// Mitsubishi GX Works2 project: 2024.06.20   PLC: Q03UDV

PROGRAM MAIN
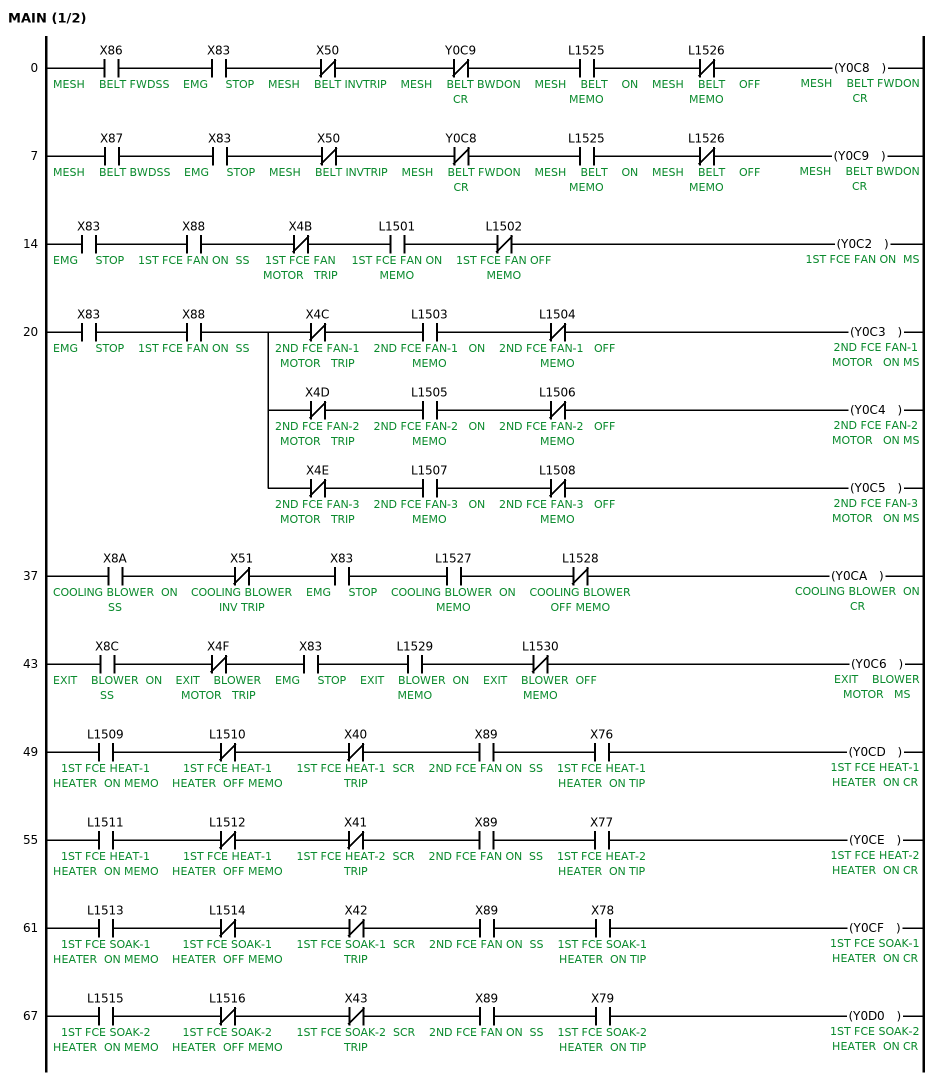
0     LD      X86  ; MESH    BELT FWDSS
      AND     X83  ; EMG     STOP
      ANI     X50  ; MESH    BELT INVTRIP
      ANI     Y0C9  ; MESH    BELT BWDON CR
      AND     L1525  ; MESH    BELT    ON MEMO
      ANI     L1526  ; MESH    BELT    OFF MEMO
      OUT     Y0C8  ; MESH    BELT FWDON CR
7     LD      X87  ; MESH    BELT BWDSS
      AND     X83  ; EMG     STOP
      ANI     X50  ; MESH    BELT INVTRIP
      ANI     Y0C8  ; MESH    BELT FWDON CR
      AND     L1525  ; MESH    BELT    ON MEMO
      ANI     L1526  ; MESH    BELT    OFF MEMO
      OUT     Y0C9  ; MESH    BELT BWDON CR
14    LD      X83  ; EMG     STOP
      AND     X88  ; 1ST FCE FAN ON  SS
      ANI     X4B  ; 1ST FCE FAN     MOTOR   TRIP
      AND     L1501  ; 1ST FCE FAN ON  MEMO
      ANI     L1502  ; 1ST FCE FAN OFF MEMO
      OUT     Y0C2  ; 1ST FCE FAN ON  MS
20    LD      X83  ; EMG     STOP
      AND     X88  ; 1ST FCE FAN ON  SS
      MPS
      ANI     X4C  ; 2ND FCE FAN-1   MOTOR   TRIP
      AND     L1503  ; 2ND FCE FAN-1   ON MEMO
      ANI     L1504  ; 2ND FCE FAN-1   OFF MEMO
      OUT     Y0C3  ; 2ND FCE FAN-1   MOTOR   ON MS
      MRD
      ANI     X4D  ; 2ND FCE FAN-2   MOTOR   TRIP
      AND     L1505  ; 2ND FCE FAN-2   ON MEMO
      ANI     L1506  ; 2ND FCE FAN-2   OFF MEMO
      OUT     Y0C4  ; 2ND FCE FAN-2   MOTOR   ON MS
      MPP
      ANI     X4E  ; 2ND FCE FAN-3   MOTOR   TRIP
      AND     L1507  ; 2ND FCE FAN-3   ON MEMO
      ANI     L1508  ; 2ND FCE FAN-3   OFF MEMO
      OUT     Y0C5  ; 2ND FCE FAN-3   MOTOR   ON MS
37    LD      X8A  ; COOLING BLOWER  ON SS
      ANI     X51  ; COOLING BLOWER  INV TRIP
      AND     X83  ; EMG     STOP
      AND     L1527  ; COOLING BLOWER  ON MEMO
      ANI     L1528  ; COOLING BLOWER  OFF MEMO
      OUT     Y0CA  ; COOLING BLOWER  ON CR
43    LD      X8C  ; EXIT    BLOWER  ON SS
      ANI     X4F  ; EXIT    BLOWER  MOTOR   TRIP
      AND     X83  ; EMG     STOP
      AND     L1529  ; EXIT    BLOWER  ON MEMO
      ANI     L1530  ; EXIT    BLOWER  OFF MEMO
      OUT     Y0C6  ; EXIT    BLOWER  MOTOR   MS
49    LD      L1509  ; 1ST FCE HEAT-1  HEATER  ON MEMO
      ANI     L1510  ; 1ST FCE HEAT-1  HEATER  OFF MEMO
      ANI     X40  ; 1ST FCE HEAT-1  SCR TRIP
      AND     X89  ; 2ND FCE FAN ON  SS
      AND     X76  ; 1ST FCE HEAT-1  HEATER  ON TIP
      OUT     Y0CD  ; 1ST FCE HEAT-1  HEATER  ON CR
55    LD      L1511  ; 1ST FCE HEAT-1  HEATER  ON MEMO
      ANI     L1512  ; 1ST FCE HEAT-1  HEATER  OFF MEMO
      ANI     X41  ; 1ST FCE HEAT-2  SCR TRIP
      AND     X89  ; 2ND FCE FAN ON  SS
      AND     X77  ; 1ST FCE HEAT-2  HEATER  ON TIP
      OUT     Y0CE  ; 1ST FCE HEAT-2  HEATER  ON CR
61    LD      L1513  ; 1ST FCE SOAK-1  HEATER  ON MEMO
      ANI     L1514  ; 1ST FCE SOAK-1  HEATER  OFF MEMO
      ANI     X42  ; 1ST FCE SOAK-1  SCR TRIP
      AND     X89  ; 2ND FCE FAN ON  SS
      AND     X78  ; 1ST FCE SOAK-1  HEATER  ON TIP
      OUT     Y0CF  ; 1ST FCE SOAK-1  HEATER  ON CR
67    LD      L1515  ; 1ST FCE SOAK-2  HEATER  ON MEMO
      ANI     L1516  ; 1ST FCE SOAK-2  HEATER  OFF MEMO
      ANI     X43  ; 1ST FCE SOAK-2  SCR TRIP
      AND     X89  ; 2ND FCE FAN ON  SS
      AND     X79  ; 1ST FCE SOAK-2  HEATER  ON TIP
      OUT     Y0D0  ; 1ST FCE SOAK-2  HEATER  ON CR
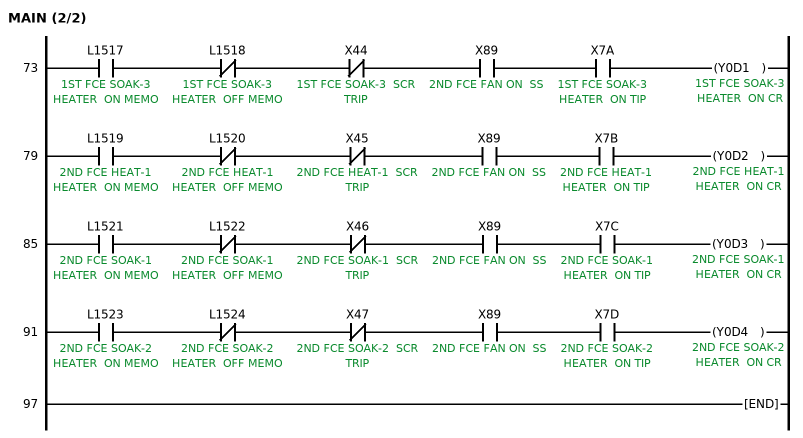
73    LD      L1517  ; 1ST FCE SOAK-3  HEATER  ON MEMO
      ANI     L1518  ; 1ST FCE SOAK-3  HEATER  OFF MEMO
      ANI     X44  ; 1ST FCE SOAK-3  SCR TRIP
      AND     X89  ; 2ND FCE FAN ON  SS
      AND     X7A  ; 1ST FCE SOAK-3  HEATER  ON TIP
      OUT     Y0D1  ; 1ST FCE SOAK-3  HEATER  ON CR
79    LD      L1519  ; 2ND FCE HEAT-1  HEATER  ON MEMO
      ANI     L1520  ; 2ND FCE HEAT-1  HEATER  OFF MEMO
      ANI     X45  ; 2ND FCE HEAT-1  SCR TRIP
      AND     X89  ; 2ND FCE FAN ON  SS
      AND     X7B  ; 2ND FCE HEAT-1  HEATER  ON TIP
      OUT     Y0D2  ; 2ND FCE HEAT-1  HEATER  ON CR
85    LD      L1521  ; 2ND FCE SOAK-1  HEATER  ON MEMO
      ANI     L1522  ; 2ND FCE SOAK-1  HEATER  OFF MEMO
      ANI     X46  ; 2ND FCE SOAK-1  SCR TRIP
      AND     X89  ; 2ND FCE FAN ON  SS
      AND     X7C  ; 2ND FCE SOAK-1  HEATER  ON TIP
      OUT     Y0D3  ; 2ND FCE SOAK-1  HEATER  ON CR
91    LD      L1523  ; 2ND FCE SOAK-2  HEATER  ON MEMO
      ANI     L1524  ; 2ND FCE SOAK-2  HEATER  OFF MEMO
      ANI     X47  ; 2ND FCE SOAK-2  SCR TRIP
      AND     X89  ; 2ND FCE FAN ON  SS
      AND     X7D  ; 2ND FCE SOAK-2  HEATER  ON TIP
      OUT     Y0D4  ; 2ND FCE SOAK-2  HEATER  ON CR
97    END
END_PROGRAM

PROGRAM HMI
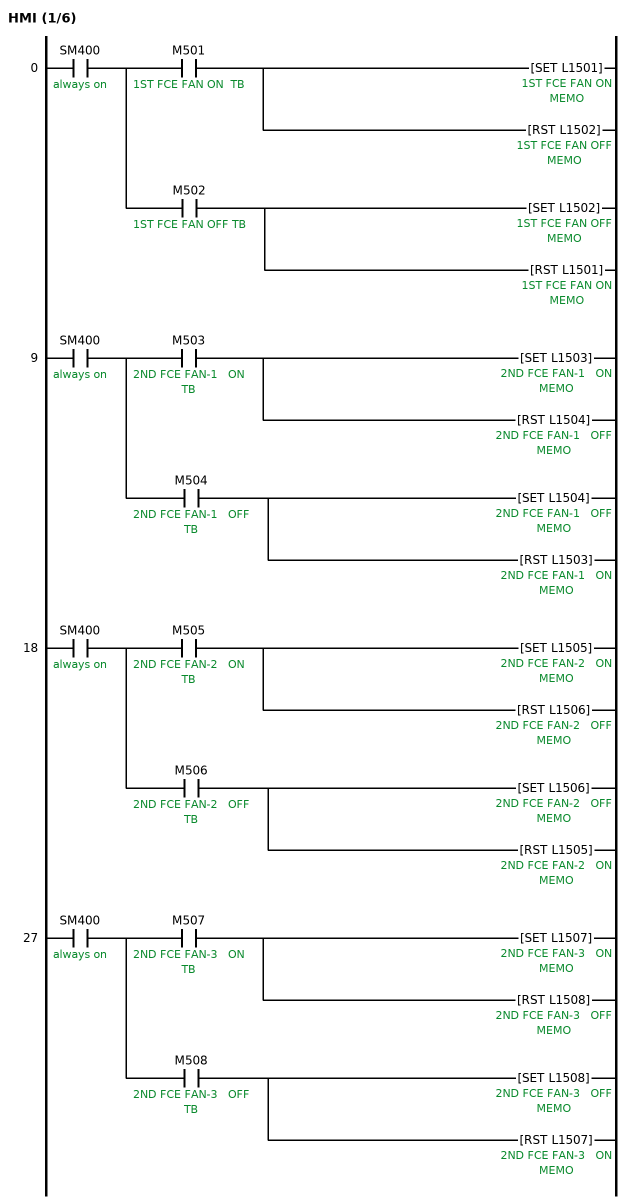
0     LD      SM400  ; always on
      MPS
      AND     M501  ; 1ST FCE FAN ON  TB
      SET     L1501  ; 1ST FCE FAN ON  MEMO
      RST     L1502  ; 1ST FCE FAN OFF MEMO
      MPP
      AND     M502  ; 1ST FCE FAN OFF TB
      SET     L1502  ; 1ST FCE FAN OFF MEMO
      RST     L1501  ; 1ST FCE FAN ON  MEMO
9     LD      SM400  ; always on
      MPS
      AND     M503  ; 2ND FCE FAN-1   ON TB
      SET     L1503  ; 2ND FCE FAN-1   ON MEMO
      RST     L1504  ; 2ND FCE FAN-1   OFF MEMO
      MPP
      AND     M504  ; 2ND FCE FAN-1   OFF TB
      SET     L1504  ; 2ND FCE FAN-1   OFF MEMO
      RST     L1503  ; 2ND FCE FAN-1   ON MEMO
18    LD      SM400  ; always on
      MPS
      AND     M505  ; 2ND FCE FAN-2   ON TB
      SET     L1505  ; 2ND FCE FAN-2   ON MEMO
      RST     L1506  ; 2ND FCE FAN-2   OFF MEMO
      MPP
      AND     M506  ; 2ND FCE FAN-2   OFF TB
      SET     L1506  ; 2ND FCE FAN-2   OFF MEMO
      RST     L1505  ; 2ND FCE FAN-2   ON MEMO
27    LD      SM400  ; always on
      MPS
      AND     M507  ; 2ND FCE FAN-3   ON TB
      SET     L1507  ; 2ND FCE FAN-3   ON MEMO
      RST     L1508  ; 2ND FCE FAN-3   OFF MEMO
      MPP
      AND     M508  ; 2ND FCE FAN-3   OFF TB
      SET     L1508  ; 2ND FCE FAN-3   OFF MEMO
      RST     L1507  ; 2ND FCE FAN-3   ON MEMO
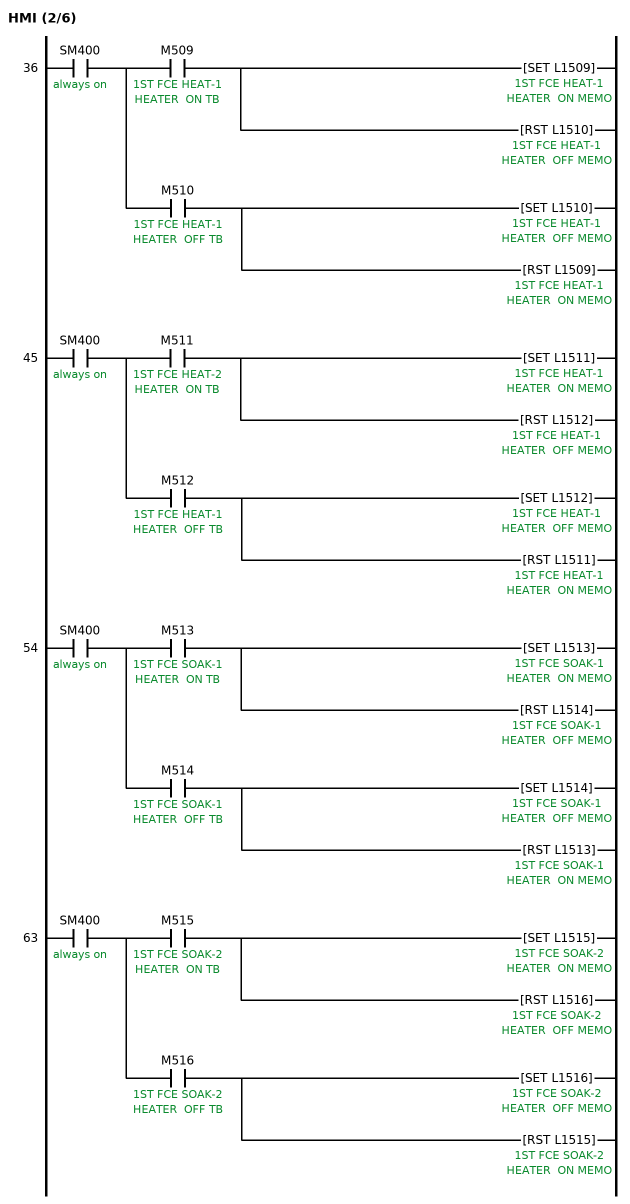
36    LD      SM400  ; always on
      MPS
      AND     M509  ; 1ST FCE HEAT-1  HEATER  ON TB
      SET     L1509  ; 1ST FCE HEAT-1  HEATER  ON MEMO
      RST     L1510  ; 1ST FCE HEAT-1  HEATER  OFF MEMO
      MPP
      AND     M510  ; 1ST FCE HEAT-1  HEATER  OFF TB
      SET     L1510  ; 1ST FCE HEAT-1  HEATER  OFF MEMO
      RST     L1509  ; 1ST FCE HEAT-1  HEATER  ON MEMO
45    LD      SM400  ; always on
      MPS
      AND     M511  ; 1ST FCE HEAT-2  HEATER  ON TB
      SET     L1511  ; 1ST FCE HEAT-1  HEATER  ON MEMO
      RST     L1512  ; 1ST FCE HEAT-1  HEATER  OFF MEMO
      MPP
      AND     M512  ; 1ST FCE HEAT-1  HEATER  OFF TB
      SET     L1512  ; 1ST FCE HEAT-1  HEATER  OFF MEMO
      RST     L1511  ; 1ST FCE HEAT-1  HEATER  ON MEMO
54    LD      SM400  ; always on
      MPS
      AND     M513  ; 1ST FCE SOAK-1  HEATER  ON TB
      SET     L1513  ; 1ST FCE SOAK-1  HEATER  ON MEMO
      RST     L1514  ; 1ST FCE SOAK-1  HEATER  OFF MEMO
      MPP
      AND     M514  ; 1ST FCE SOAK-1  HEATER  OFF TB
      SET     L1514  ; 1ST FCE SOAK-1  HEATER  OFF MEMO
      RST     L1513  ; 1ST FCE SOAK-1  HEATER  ON MEMO
63    LD      SM400  ; always on
      MPS
      AND     M515  ; 1ST FCE SOAK-2  HEATER  ON TB
      SET     L1515  ; 1ST FCE SOAK-2  HEATER  ON MEMO
      RST     L1516  ; 1ST FCE SOAK-2  HEATER  OFF MEMO
      MPP
      AND     M516  ; 1ST FCE SOAK-2  HEATER  OFF TB
      SET     L1516  ; 1ST FCE SOAK-2  HEATER  OFF MEMO
      RST     L1515  ; 1ST FCE SOAK-2  HEATER  ON MEMO
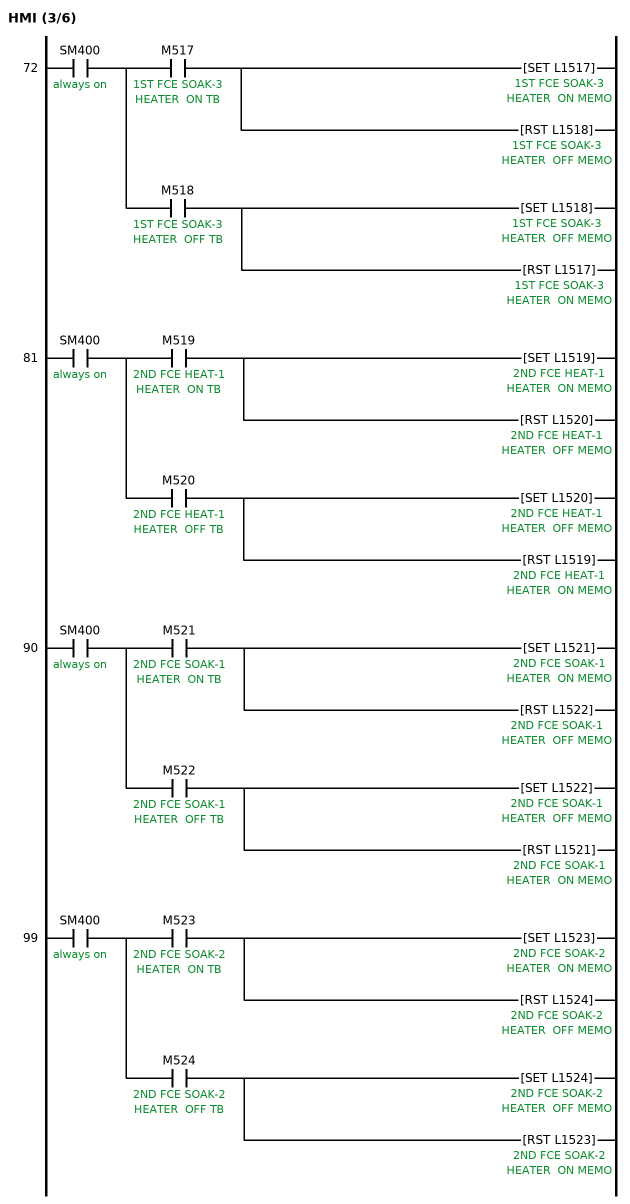
72    LD      SM400  ; always on
      MPS
      AND     M517  ; 1ST FCE SOAK-3  HEATER  ON TB
      SET     L1517  ; 1ST FCE SOAK-3  HEATER  ON MEMO
      RST     L1518  ; 1ST FCE SOAK-3  HEATER  OFF MEMO
      MPP
      AND     M518  ; 1ST FCE SOAK-3  HEATER  OFF TB
      SET     L1518  ; 1ST FCE SOAK-3  HEATER  OFF MEMO
      RST     L1517  ; 1ST FCE SOAK-3  HEATER  ON MEMO
81    LD      SM400  ; always on
      MPS
      AND     M519  ; 2ND FCE HEAT-1  HEATER  ON TB
      SET     L1519  ; 2ND FCE HEAT-1  HEATER  ON MEMO
      RST     L1520  ; 2ND FCE HEAT-1  HEATER  OFF MEMO
      MPP
      AND     M520  ; 2ND FCE HEAT-1  HEATER  OFF TB
      SET     L1520  ; 2ND FCE HEAT-1  HEATER  OFF MEMO
      RST     L1519  ; 2ND FCE HEAT-1  HEATER  ON MEMO
90    LD      SM400  ; always on
      MPS
      AND     M521  ; 2ND FCE SOAK-1  HEATER  ON TB
      SET     L1521  ; 2ND FCE SOAK-1  HEATER  ON MEMO
      RST     L1522  ; 2ND FCE SOAK-1  HEATER  OFF MEMO
      MPP
      AND     M522  ; 2ND FCE SOAK-1  HEATER  OFF TB
      SET     L1522  ; 2ND FCE SOAK-1  HEATER  OFF MEMO
      RST     L1521  ; 2ND FCE SOAK-1  HEATER  ON MEMO
99    LD      SM400  ; always on
      MPS
      AND     M523  ; 2ND FCE SOAK-2  HEATER  ON TB
      SET     L1523  ; 2ND FCE SOAK-2  HEATER  ON MEMO
      RST     L1524  ; 2ND FCE SOAK-2  HEATER  OFF MEMO
      MPP
      AND     M524  ; 2ND FCE SOAK-2  HEATER  OFF TB
      SET     L1524  ; 2ND FCE SOAK-2  HEATER  OFF MEMO
      RST     L1523  ; 2ND FCE SOAK-2  HEATER  ON MEMO
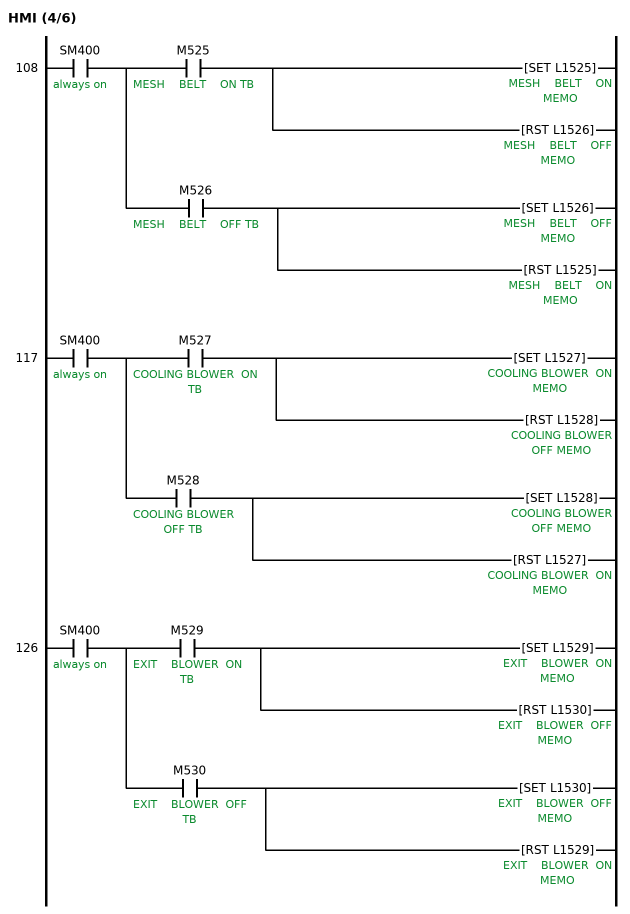
108   LD      SM400  ; always on
      MPS
      AND     M525  ; MESH    BELT    ON TB
      SET     L1525  ; MESH    BELT    ON MEMO
      RST     L1526  ; MESH    BELT    OFF MEMO
      MPP
      AND     M526  ; MESH    BELT    OFF TB
      SET     L1526  ; MESH    BELT    OFF MEMO
      RST     L1525  ; MESH    BELT    ON MEMO
117   LD      SM400  ; always on
      MPS
      AND     M527  ; COOLING BLOWER  ON TB
      SET     L1527  ; COOLING BLOWER  ON MEMO
      RST     L1528  ; COOLING BLOWER  OFF MEMO
      MPP
      AND     M528  ; COOLING BLOWER  OFF TB
      SET     L1528  ; COOLING BLOWER  OFF MEMO
      RST     L1527  ; COOLING BLOWER  ON MEMO
126   LD      SM400  ; always on
      MPS
      AND     M529  ; EXIT    BLOWER  ON TB
      SET     L1529  ; EXIT    BLOWER  ON MEMO
      RST     L1530  ; EXIT    BLOWER  OFF MEMO
      MPP
      AND     M530  ; EXIT    BLOWER  OFF TB
      SET     L1530  ; EXIT    BLOWER  OFF MEMO
      RST     L1529  ; EXIT    BLOWER  ON MEMO
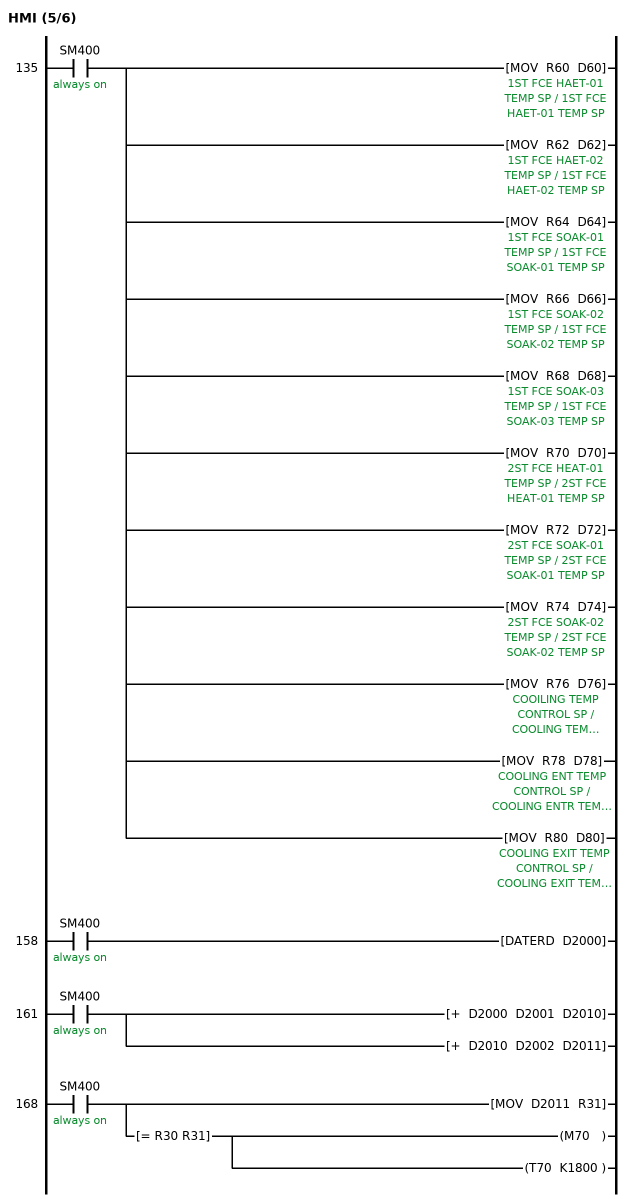
135   LD      SM400  ; always on
      MOV     R60 D60  ; 1ST FCE HAET-01 TEMP SP / 1ST FCE HAET-01 TEMP SP
      MOV     R62 D62  ; 1ST FCE HAET-02 TEMP SP / 1ST FCE HAET-02 TEMP SP
      MOV     R64 D64  ; 1ST FCE SOAK-01 TEMP SP / 1ST FCE SOAK-01 TEMP SP
      MOV     R66 D66  ; 1ST FCE SOAK-02 TEMP SP / 1ST FCE SOAK-02 TEMP SP
      MOV     R68 D68  ; 1ST FCE SOAK-03 TEMP SP / 1ST FCE SOAK-03 TEMP SP
      MOV     R70 D70  ; 2ST FCE HEAT-01 TEMP SP / 2ST FCE HEAT-01 TEMP SP
      MOV     R72 D72  ; 2ST FCE SOAK-01 TEMP SP / 2ST FCE SOAK-01 TEMP SP
      MOV     R74 D74  ; 2ST FCE SOAK-02 TEMP SP / 2ST FCE SOAK-02 TEMP SP
      MOV     R76 D76  ; COOILING TEMP CONTROL SP / COOLING TEMP CONTROL SP
      MOV     R78 D78  ; COOLING ENT TEMP CONTROL SP / COOLING ENTR TEMP CONTROL SP
      MOV     R80 D80  ; COOLING EXIT TEMP CONTROL SP / COOLING EXIT TEMP CONTROL SP
158   LD      SM400  ; always on
      DATERD  D2000
161   LD      SM400  ; always on
      +       D2000 D2001 D2010
      +       D2010 D2002 D2011
168   LD      SM400  ; always on
      MOV     D2011 R31
      AND=    R30 R31
      OUT     M70
      OUT     T70 K1800
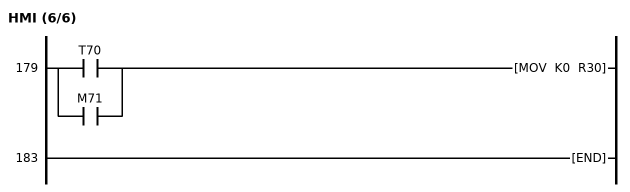
179   LD      T70
      OR      M71
      MOV     K0 R30
183   END
END_PROGRAM

PROGRAM LAMP
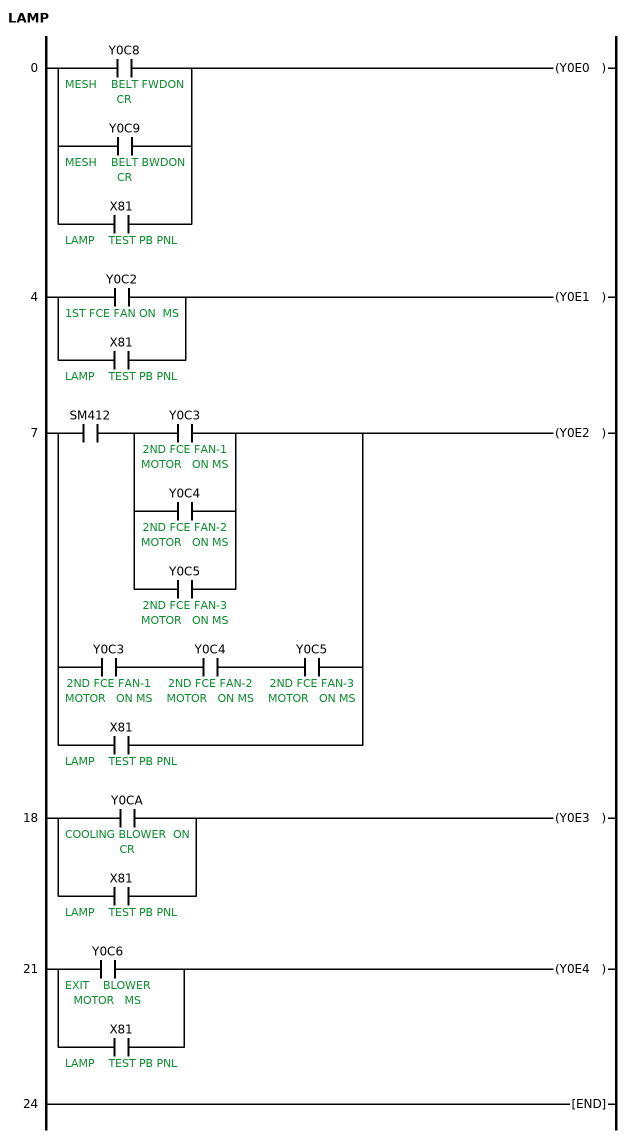
0     LD      Y0C8  ; MESH    BELT FWDON CR
      OR      Y0C9  ; MESH    BELT BWDON CR
      OR      X81  ; LAMP    TEST PB PNL
      OUT     Y0E0
4     LD      Y0C2  ; 1ST FCE FAN ON  MS
      OR      X81  ; LAMP    TEST PB PNL
      OUT     Y0E1
7     LD      SM412
      LD      Y0C3  ; 2ND FCE FAN-1   MOTOR   ON MS
      OR      Y0C4  ; 2ND FCE FAN-2   MOTOR   ON MS
      OR      Y0C5  ; 2ND FCE FAN-3   MOTOR   ON MS
      ANB
      LD      Y0C3  ; 2ND FCE FAN-1   MOTOR   ON MS
      AND     Y0C4  ; 2ND FCE FAN-2   MOTOR   ON MS
      AND     Y0C5  ; 2ND FCE FAN-3   MOTOR   ON MS
      ORB
      OR      X81  ; LAMP    TEST PB PNL
      OUT     Y0E2
18    LD      Y0CA  ; COOLING BLOWER  ON CR
      OR      X81  ; LAMP    TEST PB PNL
      OUT     Y0E3
21    LD      Y0C6  ; EXIT    BLOWER  MOTOR   MS
      OR      X81  ; LAMP    TEST PB PNL
      OUT     Y0E4
24    END
END_PROGRAM

PROGRAM ALARM
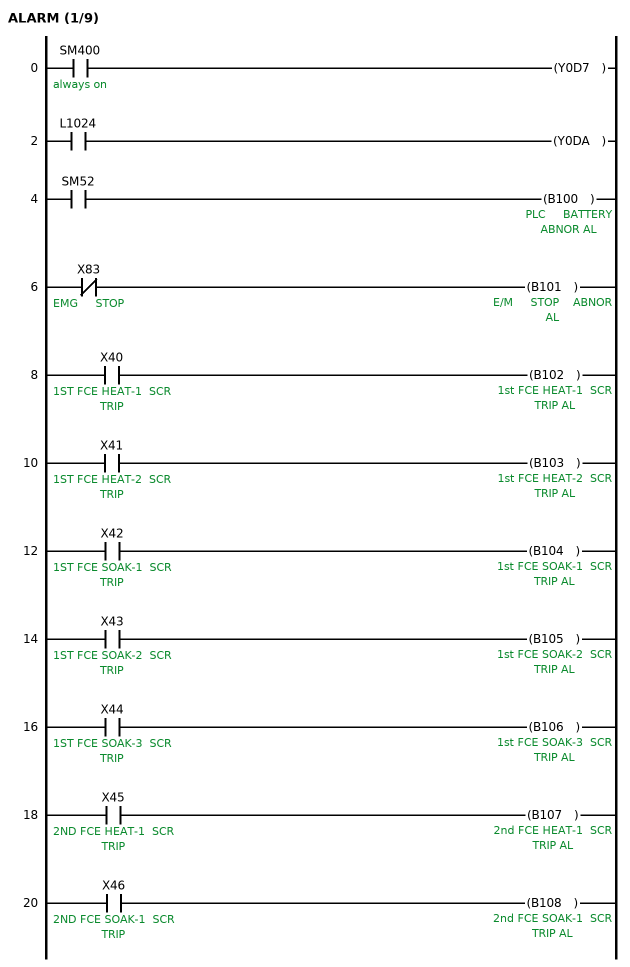
0     LD      SM400  ; always on
      OUT     Y0D7
2     LD      L1024
      OUT     Y0DA
4     LD      SM52
      OUT     B100  ; PLC     BATTERY ABNOR AL
6     LDI     X83  ; EMG     STOP
      OUT     B101  ; E/M     STOP    ABNOR AL
8     LD      X40  ; 1ST FCE HEAT-1  SCR TRIP
      OUT     B102  ; 1st FCE HEAT-1  SCR TRIP AL
10    LD      X41  ; 1ST FCE HEAT-2  SCR TRIP
      OUT     B103  ; 1st FCE HEAT-2  SCR TRIP AL
12    LD      X42  ; 1ST FCE SOAK-1  SCR TRIP
      OUT     B104  ; 1st FCE SOAK-1  SCR TRIP AL
14    LD      X43  ; 1ST FCE SOAK-2  SCR TRIP
      OUT     B105  ; 1st FCE SOAK-2  SCR TRIP AL
16    LD      X44  ; 1ST FCE SOAK-3  SCR TRIP
      OUT     B106  ; 1st FCE SOAK-3  SCR TRIP AL
18    LD      X45  ; 2ND FCE HEAT-1  SCR TRIP
      OUT     B107  ; 2nd FCE HEAT-1  SCR TRIP AL
20    LD      X46  ; 2ND FCE SOAK-1  SCR TRIP
      OUT     B108  ; 2nd FCE SOAK-1  SCR TRIP AL
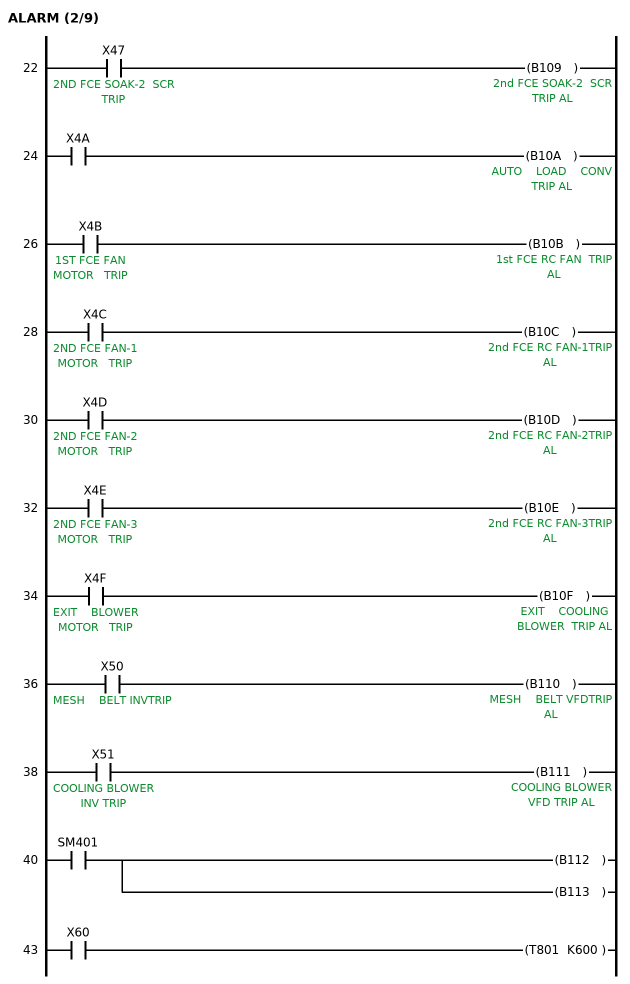
22    LD      X47  ; 2ND FCE SOAK-2  SCR TRIP
      OUT     B109  ; 2nd FCE SOAK-2  SCR TRIP AL
24    LD      X4A
      OUT     B10A  ; AUTO    LOAD    CONV    TRIP AL
26    LD      X4B  ; 1ST FCE FAN     MOTOR   TRIP
      OUT     B10B  ; 1st FCE RC FAN  TRIP AL
28    LD      X4C  ; 2ND FCE FAN-1   MOTOR   TRIP
      OUT     B10C  ; 2nd FCE RC FAN-1TRIP AL
30    LD      X4D  ; 2ND FCE FAN-2   MOTOR   TRIP
      OUT     B10D  ; 2nd FCE RC FAN-2TRIP AL
32    LD      X4E  ; 2ND FCE FAN-3   MOTOR   TRIP
      OUT     B10E  ; 2nd FCE RC FAN-3TRIP AL
34    LD      X4F  ; EXIT    BLOWER  MOTOR   TRIP
      OUT     B10F  ; EXIT    COOLING BLOWER  TRIP AL
36    LD      X50  ; MESH    BELT INVTRIP
      OUT     B110  ; MESH    BELT VFDTRIP AL
38    LD      X51  ; COOLING BLOWER  INV TRIP
      OUT     B111  ; COOLING BLOWER  VFD TRIP AL
40    LD      SM401
      OUT     B112
      OUT     B113
43    LD      X60
      OUT     T801 K600
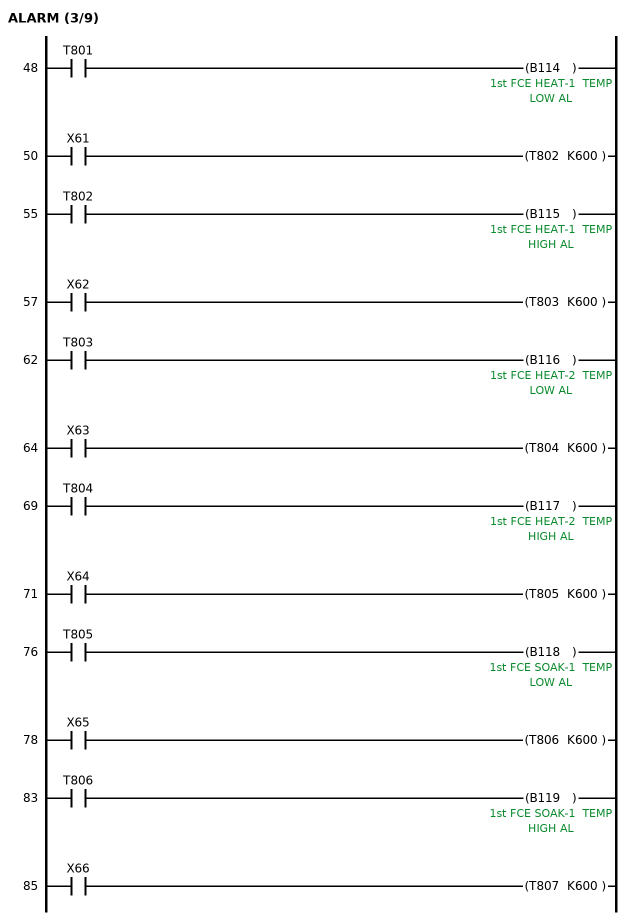
48    LD      T801
      OUT     B114  ; 1st FCE HEAT-1  TEMP    LOW AL
50    LD      X61
      OUT     T802 K600
55    LD      T802
      OUT     B115  ; 1st FCE HEAT-1  TEMP    HIGH AL
57    LD      X62
      OUT     T803 K600
62    LD      T803
      OUT     B116  ; 1st FCE HEAT-2  TEMP    LOW AL
64    LD      X63
      OUT     T804 K600
69    LD      T804
      OUT     B117  ; 1st FCE HEAT-2  TEMP    HIGH AL
71    LD      X64
      OUT     T805 K600
76    LD      T805
      OUT     B118  ; 1st FCE SOAK-1  TEMP    LOW AL
78    LD      X65
      OUT     T806 K600
83    LD      T806
      OUT     B119  ; 1st FCE SOAK-1  TEMP    HIGH AL
85    LD      X66
      OUT     T807 K600
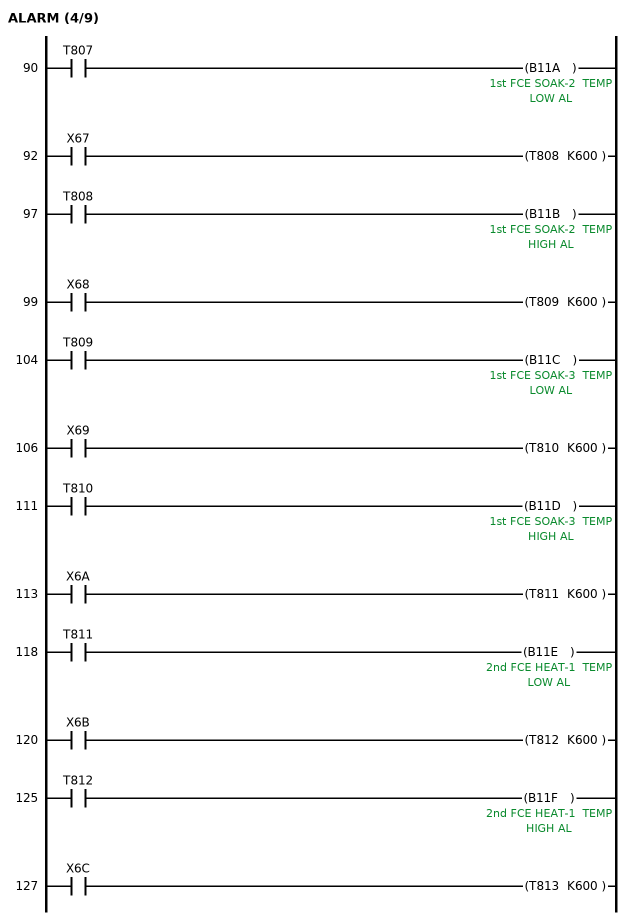
90    LD      T807
      OUT     B11A  ; 1st FCE SOAK-2  TEMP    LOW AL
92    LD      X67
      OUT     T808 K600
97    LD      T808
      OUT     B11B  ; 1st FCE SOAK-2  TEMP    HIGH AL
99    LD      X68
      OUT     T809 K600
104   LD      T809
      OUT     B11C  ; 1st FCE SOAK-3  TEMP    LOW AL
106   LD      X69
      OUT     T810 K600
111   LD      T810
      OUT     B11D  ; 1st FCE SOAK-3  TEMP    HIGH AL
113   LD      X6A
      OUT     T811 K600
118   LD      T811
      OUT     B11E  ; 2nd FCE HEAT-1  TEMP    LOW AL
120   LD      X6B
      OUT     T812 K600
125   LD      T812
      OUT     B11F  ; 2nd FCE HEAT-1  TEMP    HIGH AL
127   LD      X6C
      OUT     T813 K600
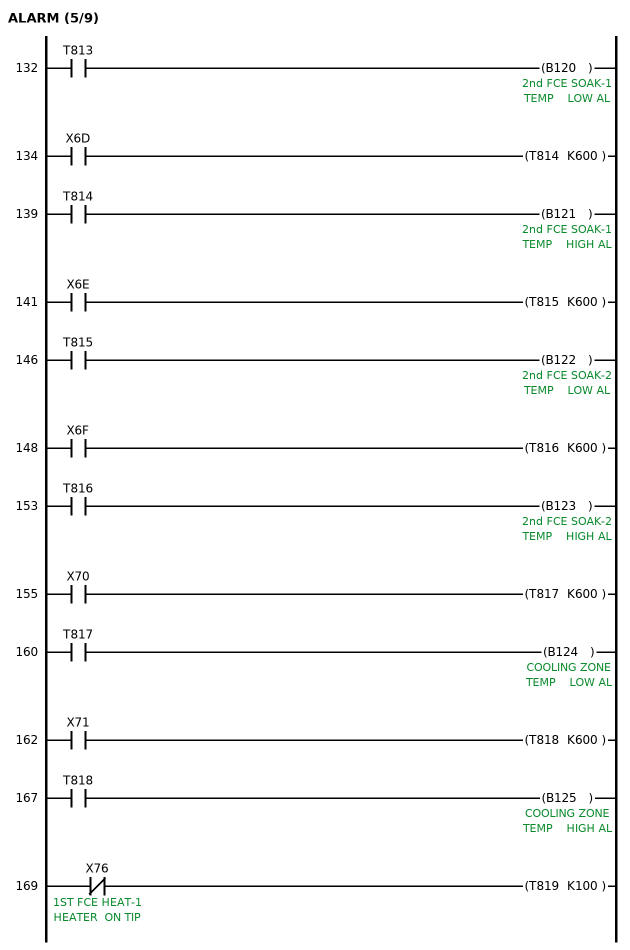
132   LD      T813
      OUT     B120  ; 2nd FCE SOAK-1  TEMP    LOW AL
134   LD      X6D
      OUT     T814 K600
139   LD      T814
      OUT     B121  ; 2nd FCE SOAK-1  TEMP    HIGH AL
141   LD      X6E
      OUT     T815 K600
146   LD      T815
      OUT     B122  ; 2nd FCE SOAK-2  TEMP    LOW AL
148   LD      X6F
      OUT     T816 K600
153   LD      T816
      OUT     B123  ; 2nd FCE SOAK-2  TEMP    HIGH AL
155   LD      X70
      OUT     T817 K600
160   LD      T817
      OUT     B124  ; COOLING ZONE    TEMP    LOW AL
162   LD      X71
      OUT     T818 K600
167   LD      T818
      OUT     B125  ; COOLING ZONE    TEMP    HIGH AL
169   LDI     X76  ; 1ST FCE HEAT-1  HEATER  ON TIP
      OUT     T819 K100
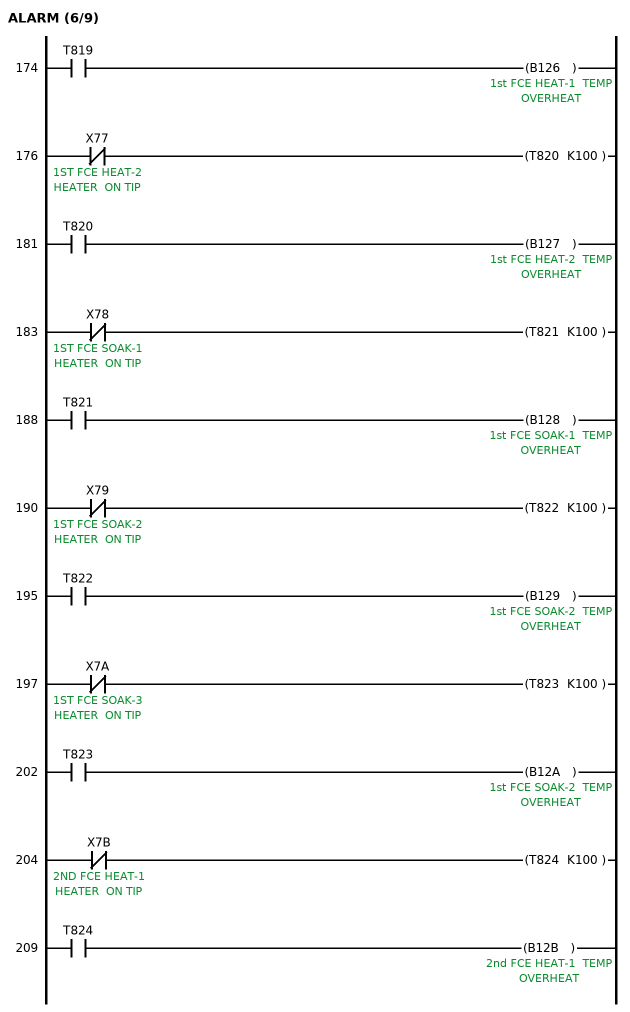
174   LD      T819
      OUT     B126  ; 1st FCE HEAT-1  TEMP    OVERHEAT
176   LDI     X77  ; 1ST FCE HEAT-2  HEATER  ON TIP
      OUT     T820 K100
181   LD      T820
      OUT     B127  ; 1st FCE HEAT-2  TEMP    OVERHEAT
183   LDI     X78  ; 1ST FCE SOAK-1  HEATER  ON TIP
      OUT     T821 K100
188   LD      T821
      OUT     B128  ; 1st FCE SOAK-1  TEMP    OVERHEAT
190   LDI     X79  ; 1ST FCE SOAK-2  HEATER  ON TIP
      OUT     T822 K100
195   LD      T822
      OUT     B129  ; 1st FCE SOAK-2  TEMP    OVERHEAT
197   LDI     X7A  ; 1ST FCE SOAK-3  HEATER  ON TIP
      OUT     T823 K100
202   LD      T823
      OUT     B12A  ; 1st FCE SOAK-2  TEMP    OVERHEAT
204   LDI     X7B  ; 2ND FCE HEAT-1  HEATER  ON TIP
      OUT     T824 K100
209   LD      T824
      OUT     B12B  ; 2nd FCE HEAT-1  TEMP    OVERHEAT
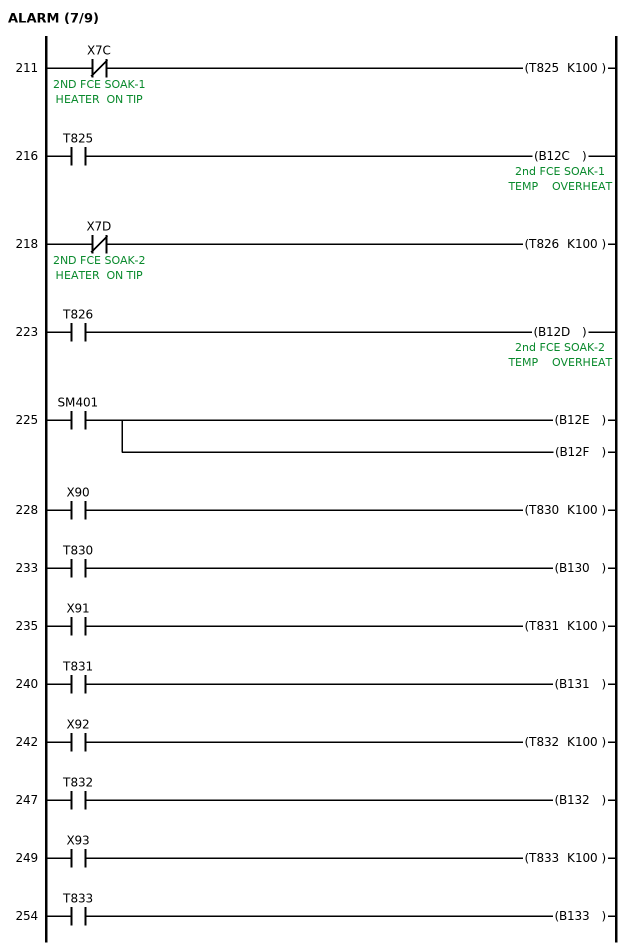
211   LDI     X7C  ; 2ND FCE SOAK-1  HEATER  ON TIP
      OUT     T825 K100
216   LD      T825
      OUT     B12C  ; 2nd FCE SOAK-1  TEMP    OVERHEAT
218   LDI     X7D  ; 2ND FCE SOAK-2  HEATER  ON TIP
      OUT     T826 K100
223   LD      T826
      OUT     B12D  ; 2nd FCE SOAK-2  TEMP    OVERHEAT
225   LD      SM401
      OUT     B12E
      OUT     B12F
228   LD      X90
      OUT     T830 K100
233   LD      T830
      OUT     B130
235   LD      X91
      OUT     T831 K100
240   LD      T831
      OUT     B131
242   LD      X92
      OUT     T832 K100
247   LD      T832
      OUT     B132
249   LD      X93
      OUT     T833 K100
254   LD      T833
      OUT     B133
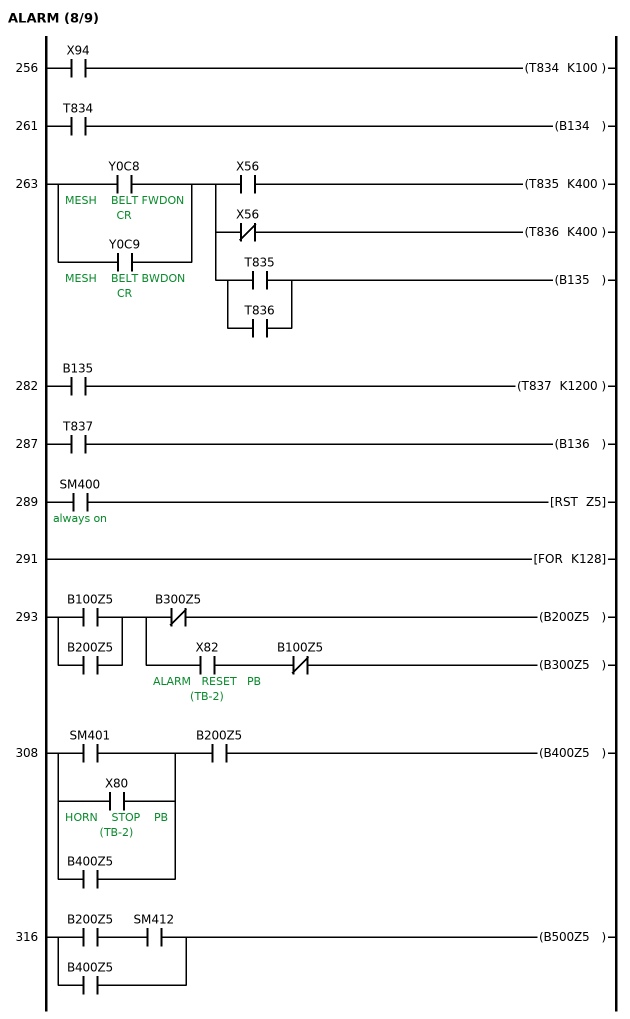
256   LD      X94
      OUT     T834 K100
261   LD      T834
      OUT     B134
263   LD      Y0C8  ; MESH    BELT FWDON CR
      OR      Y0C9  ; MESH    BELT BWDON CR
      MPS
      AND     X56
      OUT     T835 K400
      MRD
      ANI     X56
      OUT     T836 K400
      MPP
      LD      T835
      OR      T836
      ANB
      OUT     B135
282   LD      B135
      OUT     T837 K1200
287   LD      T837
      OUT     B136
289   LD      SM400  ; always on
      RST     Z5
291   FOR     K128
293   LD      B100Z5
      OR      B200Z5
      MPS
      ANI     B300Z5
      OUT     B200Z5
      MPP
      AND     X82  ; ALARM   RESET   PB      (TB-2)
      ANI     B100Z5
      OUT     B300Z5
308   LD      SM401
      OR      X80  ; HORN    STOP    PB      (TB-2)
      OR      B400Z5
      AND     B200Z5
      OUT     B400Z5
316   LD      B200Z5
      AND     SM412
      OR      B400Z5
      OUT     B500Z5
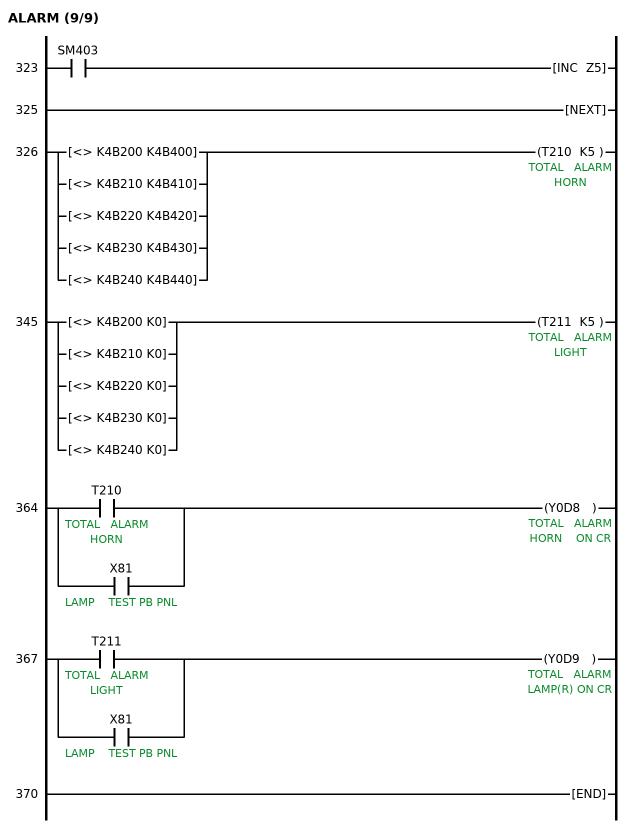
323   LD      SM403
      INC     Z5
325   NEXT
326   LD<>    K4B200 K4B400
      OR<>    K4B210 K4B410
      OR<>    K4B220 K4B420
      OR<>    K4B230 K4B430
      OR<>    K4B240 K4B440
      OUT     T210 K5  ; TOTAL   ALARM   HORN
345   LD<>    K4B200 K0
      OR<>    K4B210 K0
      OR<>    K4B220 K0
      OR<>    K4B230 K0
      OR<>    K4B240 K0
      OUT     T211 K5  ; TOTAL   ALARM   LIGHT
364   LD      T210  ; TOTAL   ALARM   HORN
      OR      X81  ; LAMP    TEST PB PNL
      OUT     Y0D8  ; TOTAL   ALARM   HORN    ON CR
367   LD      T211  ; TOTAL   ALARM   LIGHT
      OR      X81  ; LAMP    TEST PB PNL
      OUT     Y0D9  ; TOTAL   ALARM   LAMP(R) ON CR
370   END
END_PROGRAM

PROGRAM COMMUN
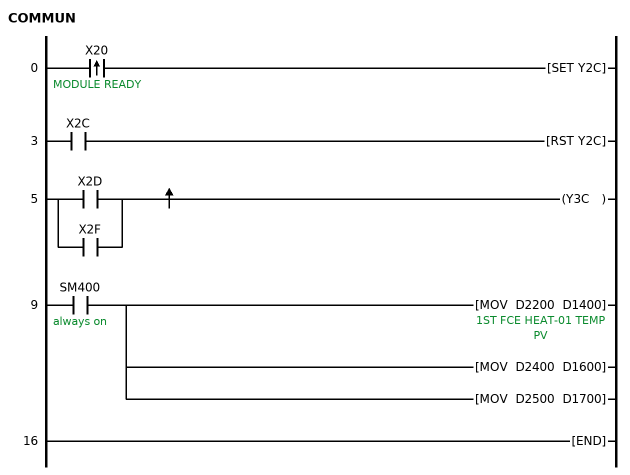
0     LDP     X20  ; MODULE READY
      SET     Y2C
3     LD      X2C
      RST     Y2C
5     LD      X2D
      OR      X2F
      MEP
      OUT     Y3C
9     LD      SM400  ; always on
      MOV     D2200 D1400  ; 1ST FCE HEAT-01 TEMP PV
      MOV     D2400 D1600
      MOV     D2500 D1700
16    END
END_PROGRAM

PROGRAM COMMUNIC
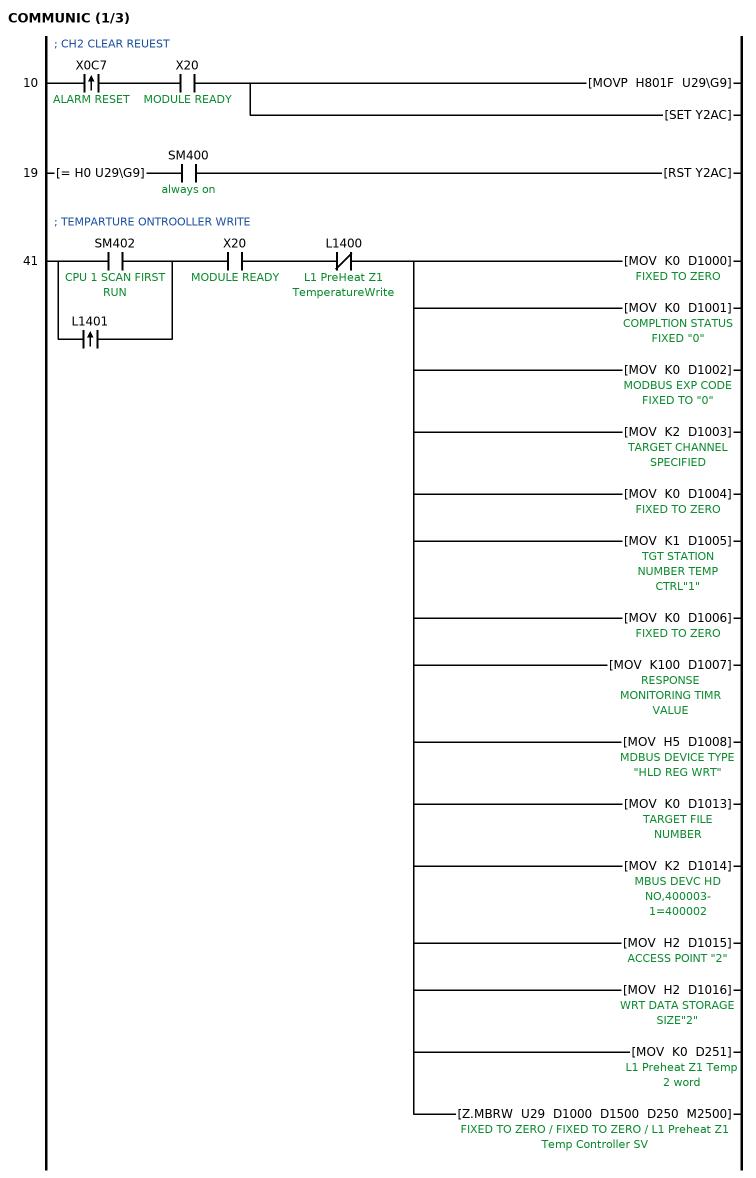
; CH2 CLEAR REUEST
10    LDP     X0C7  ; ALARM RESET
      AND     X20  ; MODULE READY
      MOVP    H801F U29\G9
      SET     Y2AC
19    LD=     H0 U29\G9
      AND     SM400  ; always on
      RST     Y2AC
; TEMPARTURE ONTROOLLER WRITE
41    LD      SM402  ; CPU 1 SCAN FIRST RUN
      ORP     L1401
      AND     X20  ; MODULE READY
      ANI     L1400  ; L1 PreHeat Z1 TemperatureWrite
      MOV     K0 D1000  ; FIXED TO ZERO
      MOV     K0 D1001  ; COMPLTION STATUS FIXED "0"
      MOV     K0 D1002  ; MODBUS EXP CODE FIXED TO "0"
      MOV     K2 D1003  ; TARGET CHANNEL SPECIFIED
      MOV     K0 D1004  ; FIXED TO ZERO
      MOV     K1 D1005  ; TGT STATION NUMBER TEMP CTRL"1"
      MOV     K0 D1006  ; FIXED TO ZERO
      MOV     K100 D1007  ; RESPONSE MONITORING TIMR VALUE
      MOV     H5 D1008  ; MDBUS DEVICE TYPE "HLD REG WRT"
      MOV     K0 D1013  ; TARGET FILE NUMBER
      MOV     K2 D1014  ; MBUS DEVC HD NO,400003-1=400002
      MOV     H2 D1015  ; ACCESS POINT "2"
      MOV     H2 D1016  ; WRT DATA STORAGE SIZE"2"
      MOV     K0 D251  ; L1 Preheat Z1 Temp 2 word
      Z.MBRW  U29 D1000 D1500 D250 M2500  ; FIXED TO ZERO / L1 Preheat Z1 Temp Controller SV
        [note] MODBUS READ/WRITE INSTRUCTION
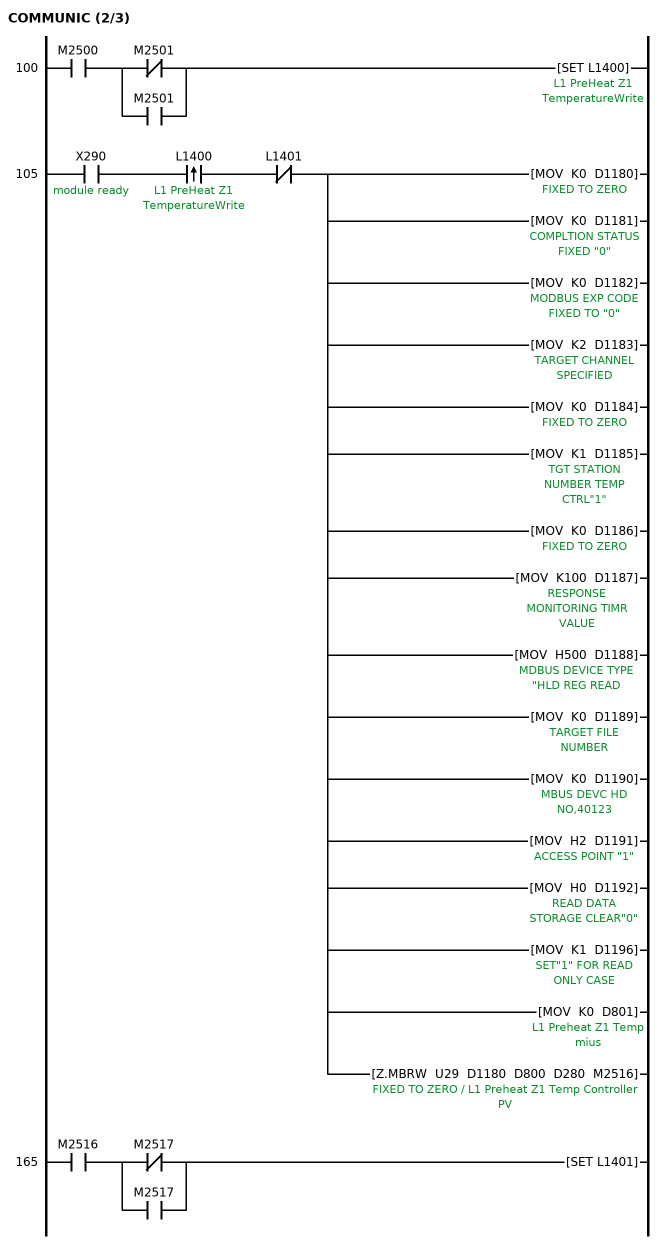
100   LD      M2500
      LDI     M2501
      OR      M2501
      ANB
      SET     L1400  ; L1 PreHeat Z1 TemperatureWrite
105   LD      X290  ; module ready
      ANDP    L1400  ; L1 PreHeat Z1 TemperatureWrite
      ANI     L1401
      MOV     K0 D1180  ; FIXED TO ZERO
      MOV     K0 D1181  ; COMPLTION STATUS FIXED "0"
      MOV     K0 D1182  ; MODBUS EXP CODE FIXED TO "0"
      MOV     K2 D1183  ; TARGET CHANNEL SPECIFIED
      MOV     K0 D1184  ; FIXED TO ZERO
      MOV     K1 D1185  ; TGT STATION NUMBER TEMP CTRL"1"
      MOV     K0 D1186  ; FIXED TO ZERO
      MOV     K100 D1187  ; RESPONSE MONITORING TIMR VALUE
      MOV     H500 D1188  ; MDBUS DEVICE TYPE "HLD REG READ
      MOV     K0 D1189  ; TARGET FILE NUMBER
      MOV     K0 D1190  ; MBUS DEVC HD NO,40123
      MOV     H2 D1191  ; ACCESS POINT "1"
      MOV     H0 D1192  ; READ DATA STORAGE CLEAR"0"
      MOV     K1 D1196  ; SET"1" FOR READ ONLY CASE
      MOV     K0 D801  ; L1 Preheat Z1 Temp mius
      Z.MBRW  U29 D1180 D800 D280 M2516  ; L1 Preheat Z1 Temp Controller PV
        [note] MODBUS READ/WRITE INSTRUCTION
165   LD      M2516
      LDI     M2517
      OR      M2517
      ANB
      SET     L1401
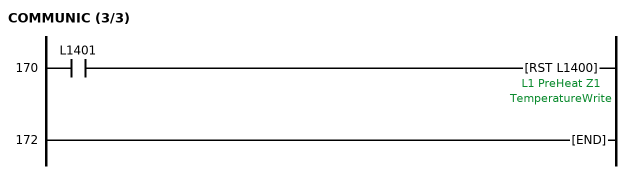
170   LD      L1401
      RST     L1400  ; L1 PreHeat Z1 TemperatureWrite
172   END
END_PROGRAM

// device comments not shown above
X0  ; MODULE READY
X10  ; INTELGENT FU CTION MODULE SETTIN
Y0BC  ; CH2 ERROE CLEAR REQUEST
L1431  ; REPEAT CYCLE
D201  ; COMPLTION STATUS FIXED "0"
D202  ; MODBUS EXP CODE FIXED TO "0"
D203  ; TARGET CHANNEL SPECIFIED
D205  ; TGT STATION NUMBER TEMP CTRL"1"
D207  ; RESPONSE MONITORING TIMR VALUE
D208  ; MDBUS DEVICE TYPE "HLD REG WRT"
D209  ; READ AREA ZERO
D210  ; MODBUS WRITE ADD 40003
D211  ; READ AREA ZERO
D212  ; READ DATR STORAGE
D213  ; TARGET FILE NUMBER
D214  ; MBUS DEVC ADDRE 40001
D215  ; ACCESS POINT "1"
D216  ; WRT DATA STORAGE SIZE"1"
D2100  ; 1ST FCE HEAT-01 TEMP PV
D2101  ; 1ST FCE HEAT-02 TEMP PV
D2102  ; 1ST FCE SOAK-01 TEMP PV
D2103  ; 1ST FCE SOAK-02 TEMP PV
D2104  ; 1ST FCE SOAK-03 TEMP PV
D2105  ; 2ST FCE HEAT-01 TEMP PV
D2106  ; 2ST FCE SOAK-01 TEMP PV
D2107  ; 2ST FCE SOAK-02 TEMP PV
D2108  ; COOLING TEMP CONTROL
D2109  ; COOLING ENTRAN TEMP CONTROL PV
D2110  ; COOLING EXIT TEMP CONTROL PV
D2111  ; MESH BELT MOTOR HZ PV
D2201  ; 1ST FCE HEAT-02 TEMP PV
D2202  ; 1ST FCE SOAK-01 TEMP PV
D2203  ; 1ST FCE SOAK-02 TEMP PV
D2204  ; 1ST FCE SOAK-03 TEMP PV
D2205  ; 2ST FCE HEAT-01 TEMP PV
D2206  ; 2ST FCE SOAK-01 TEMP PV
D2207  ; 2ST FCE SOAK-02 TEMP PV
D2208  ; COOLING TEMP CONTROL
D2209  ; COOLING ENTRAN TEMP CONTROL PV
D2210  ; COOLING EXIT TEMP CONTROL PV
D2211  ; MESH BELT MOTOR HZ PV
